(* IEC 61131-3 sources: SortJet_MasterSPS_Aufbau.fbsproj/09_Station/Shuttle/[101,102] Shuttle/Aktionen, 4 files *)

(* ---- Shuttle_Ansteuerung_Ressourcen_FB_V01_00_00.fb.st ---- *)
(* METADATA
{
	"v3Meta": {
		"objectGuid": "9404f6fa-2a6f-44db-8f42-3f6f32f76ed1"
	}
}
*)
FUNCTION_BLOCK Shuttle_Ansteuerung_Ressourcen_FB_V01_00_00 EXTENDS Basic_Shuttle_Aktion_FB_V01_00_00
VAR_INPUT

  // GREIFER [Ausbaustufe stStationsAufbau.bGreifer]
  bpGreiferAktiv : BOOL;
  Greifer        : REFERENCE TO Shuttle_Greifer_FB_V01_00_00;

END_VAR
VAR
  tonlTimeout : TON;

  // BOOL
  blMitGreifer : BOOL; // Vorab-Auftrag mit Greiferseite und Greifer vorhanden
  blGlasUeberspringen : BOOL; // Vorab ohne Glasaktion: Eintransport aktiv oder gerade gewesen
END_VAR
//-------------------------------------------------------------------------------------------------
// AKTION ANSTEUERUNG RESOURCEN WAEHREND DER QUERFAHRT
//-------------------------------------------------------------------------------------------------
(* Wichtig:
   - Es handelt isch hier um eine Aktion die waehrend der Shuttlequerfahrt [Verfahrauftrag] abgearbeitet wird.
   - Zu beachten ist das:
     => Wenn der Riemen verfahrern werden soll pruefen ob der autarke Vortransport aktiv ist
     => Aktion laeuft parallel zum Verfahrauftrag der Oberflaeche
*)
IF (  BasisStationsParameter.bVorabKomponentenAnsteuerung[wWand]
     AND bpAutomatikAktiv )
THEN

  // Ausnahmesituation
  IF ( Glastransport.bpFehler ) THEN
    Glastransport.bpVortransport              := FALSE;
    Glastransport.bpVortransportRueck         := FALSE;
    Glastransport.bpStarteVorabPositionierung := FALSE;
    Glastransport.bpStarteVorabPositionierungRueckwaertig := FALSE;
    BasisStationsParameter.wFehlerNummer := Glastransport.wpFehlerNr;
    steplAktion := STEP_900_E;
  END_IF

  IF ( Kippen.bpFehler ) THEN
    Kippen.bpPositionieren := FALSE;
    BasisStationsParameter.wFehlerNummer :=  Kippen.wpFehlerNr;
    steplAktion := STEP_900_E;
  END_IF

  IF ( Wandverstellung.bpFehler ) THEN
    Wandverstellung.bpStartePositionierung := FALSE;
    BasisStationsParameter.wFehlerNummer :=  Wandverstellung.wpFehlerNr;
    steplAktion := STEP_900_E;
  END_IF

  IF ( blMitGreifer AND Greifer.bpFehler ) THEN
    Greifer.bpPositionieren                         := FALSE;
    Greifer.bpStarteVorabPositionierungEintransport := FALSE;
    BasisStationsParameter.awFehlerInformationen    := Greifer.awpFehlerInformationen;
    BasisStationsParameter.awFehlerInformationen[1] := Greifer.wpFehlerKennung;
    BasisStationsParameter.wFehlerNummer            := Greifer.wpFehlerNr;
    steplAktion := STEP_900_E;
  END_IF

  (* Hinweis:
     - Starten der Schrittkette
  *)
  CASE steplAktion OF
    // VORAB KOMPONENTEN ANSTEUERUNG ========================
    STEP_0_E:
      BasisStationsParameter.bVorabKomponentenAnsteuerungAbgeschlossen[wWand] := FALSE;
      tonlTimeout( IN := FALSE );

      blMitGreifer :=     bpGreiferAktiv
                      AND ( BasisStationsParameter.pVorAbAuftragsdaten[wWand].stAuftragsOptionen.eGreiferTyp <> eGreiferDefault );

      IF ( BasisStationsParameter.stMKs.stStationsOptionen.bVorAbKomponentenAnsteuerung ) THEN
        steplAktion := STEP_10_E;
      ELSE
        steplAktion := STEP_1000_E;
      END_IF

    // VORAB KOMPONENTEN ANSTEUERUNG WAND 1 ========================
    STEP_10_E:
      (* Hinweis:
         - Wandverstellung ansteuern
         - Kippen ansteuern
         - Erst wenn der Glastransport seinen Eintransport beendet hat: Ein vorzeitig quittierter
           Eintransport (letzte Scheibe, Freigabe Querfahrt) laeuft im Glastransport noch weiter,
           waehrend bEintransport bereits FALSE ist. Kippen, Wandverstellung und Greifer duerfen
           die noch fahrende Scheibe nicht beeinflussen (Fehler: Scheibe faehrt auf den Auslaufstopp).
      *)
      IF (     NOT Glastransport.bpEintransport
           AND NOT Glastransport.bpRueckwaertsEintransportieren )
      THEN
        Wandverstellung.epSollStellung         := BasisStationsParameter.pVorAbAuftragsdaten[wWand].stAuftragsOptionen.eDickenverstellung;
        Wandverstellung.bpStartePositionierung := TRUE;

        IF BasisStationsParameter.pVorAbAuftragsdaten[wWand].stAuftragsOptionen.eKippen_SollPosition <> eKippen_Default THEN
          Kippen.epZielPosition := BasisStationsParameter.pVorAbAuftragsdaten[wWand].stAuftragsOptionen.eKippen_SollPosition;
          Kippen.bpPositionieren := TRUE;
        END_IF

        steplAktion := STEP_20_E;
      END_IF

    // VORAB KOMPONENTEN ANSTEUERUNG WAND 1 ========================
    STEP_20_E:
      (* Hinweis:
         - Glastransport ansteuern
         - Laeuft der Eintransport noch (bEintransport) oder ist er gerade abgeschlossen (Eintransport gewesen),
           liegt die Scheibe definiert: die Glasaktion der Vorab entfaellt, es wird nicht gewartet
         - Jede weitere Vorab positioniert die Scheibe neu (Sensor erst freifahren, dann neu anfahren)
      *)
      blGlasUeberspringen := BasisStationsParameter.bEintransport[wWand]
                             OR BasisStationsParameter.bEintransportGewesen[wWand];
      BasisStationsParameter.bEintransportGewesen[wWand] := FALSE;

      IF ( NOT blGlasUeberspringen
           AND NOT Glastransport.bpEintransport
           AND NOT Glastransport.bpRueckwaertsEintransportieren )
      THEN

        CASE BasisStationsParameter.pVorAbAuftragsdaten[wWand].stAuftragsOptionen.eGlastransport OF

          eGlastransport_Default:
            ;

          eGlastransport_AufEinlauf:
            Glastransport.bpStarteVorabPositionierungRueckwaertig := NOT Glastransport.bpAuftragAktiv;

          eGlastransport_AufEinlaufVorab:
            Glastransport.bpVortransportRueck := TRUE;

          eGlastransport_AufAuslauf,
            eGlastransport_AufAuslaufVorab:
            Glastransport.bpStarteVorabPositionierung := NOT Glastransport.bpAuftragAktiv;

        END_CASE

      END_IF

      (* Hinweis:
         - Greifer [Ausbaustufe] waehrend der Querfahrt vorpositionieren
           => Austransport: Greifer hinter die Glaskante stellen
           => Eintransport: Greifer an die Wandseite stellen und ausfahren
         - Entfaellt solange der Eintransport noch aktiv ist (Auftrag oder Glastransport)
      *)
      IF (     blMitGreifer
           AND NOT Greifer.bpAuftragAktiv
           AND NOT BasisStationsParameter.bEintransport[wWand]
           AND NOT Glastransport.bpEintransport
           AND NOT Glastransport.bpRueckwaertsEintransportieren )
      THEN
        Greifer.epGreiferTyp := BasisStationsParameter.pVorAbAuftragsdaten[wWand].stAuftragsOptionen.eGreiferTyp;

        IF ( BasisStationsParameter.pVorAbAuftragsdaten[wWand].wAuftragstyp.0 ) THEN
          Greifer.rpGlaslaenge    := BasisStationsParameter.pVorAbAuftragsdaten[wWand].rLaenge;
          Greifer.bpPositionieren := TRUE;
        ELSE
          Greifer.bpStarteVorabPositionierungEintransport := NOT Greifer.bpVorpositioniertEintransport;
        END_IF
      END_IF

      tonlTimeout( IN := FALSE );
      steplAktion := STEP_100_E;

    // VORAB KOMPONENTEN ANSTEUERUNG WAND 1 ========================
    STEP_100_E:
      (* Hinweis:
         - Einsammeln aller ausgelösten Ereignisse auf bpDone
      *)
      // Nach 60s Fehler melden, dass die Komponenten nicht fertig werden
      tonlTimeout(IN := TRUE, PT := T#60S);

      IF (   ( Kippen.bpDone OR NOT Kippen.bpPositionieren )
           AND (( Glastransport.bpVortransport AND Glastransport.bpDone) OR NOT Glastransport.bpVortransport)
           AND (( Glastransport.bpVortransportRueck AND Glastransport.bpDone) OR NOT Glastransport.bpVortransportRueck)
           AND (( Glastransport.bpStarteVorabPositionierung AND Glastransport.bpDone) OR NOT Glastransport.bpStarteVorabPositionierung)
           AND (( Glastransport.bpStarteVorabPositionierungRueckwaertig AND Glastransport.bpDone) OR NOT Glastransport.bpStarteVorabPositionierungRueckwaertig)
           AND (( Wandverstellung.bpStartePositionierung AND Wandverstellung.bpDone) OR NOT Wandverstellung.bpStartePositionierung)
           AND (    NOT blMitGreifer
                 OR (     (( Greifer.bpPositionieren AND Greifer.bpPositionierungAbgeschlossen ) OR NOT Greifer.bpPositionieren )
                      AND (( Greifer.bpStarteVorabPositionierungEintransport AND Greifer.bpVorabPositionierungEintransportAbgeschlossen ) OR NOT Greifer.bpStarteVorabPositionierungEintransport ) ) ) )
      THEN

        Glastransport.bpVortransport                    := FALSE;
        Glastransport.bpVortransportRueck               := FALSE;
        Glastransport.bpStarteVorabPositionierung       := FALSE;
        Glastransport.bpStarteVorabPositionierungRueckwaertig := FALSE;

        Wandverstellung.bpStartePositionierung          := FALSE;
        Kippen.bpPositionieren                          := FALSE;

        IF ( blMitGreifer ) THEN
          Greifer.bpPositionieren                         := FALSE;
          Greifer.bpStarteVorabPositionierungEintransport := FALSE;
        END_IF

        steplAktion := STEP_1000_E;
      END_IF

      IF tonlTimeout.Q THEN
        BasisStationsParameter.wFehlerNummer := cMELDUNG_STATION_VORABKOMPONENTENANSTEUERUN_NOT_DONE;
        steplAktion := STEP_900_E;
      END_IF

    // VORAB KOMPONENTEN ANSTEUERUNG WAND 1 ========================
    STEP_900_E:
      BasisStationsParameter.bFehler := TRUE;

    // VORAB KOMPONENTEN ANSTEUERUNG WAND 1 ========================
    STEP_1000_E:

      Glastransport.bpVortransport                    := FALSE;
      Glastransport.bpVortransportRueck               := FALSE;
      Glastransport.bpStarteVorabPositionierung       := FALSE;
      Glastransport.bpStarteVorabPositionierungRueckwaertig := FALSE;

      Wandverstellung.bpStartePositionierung          := FALSE;
      Kippen.bpPositionieren                          := FALSE;

      BasisStationsParameter.bVorabKomponentenAnsteuerungAbgeschlossen[wWand] := TRUE;

  // VORAB KOMPONENTEN ANSTEUERUNG WAND 1 ========================
  END_CASE

END_IF

IF ( NOT BasisStationsParameter.bVorabKomponentenAnsteuerung[wWand] ) THEN

  IF ( steplAktion > STEP_0_E ) THEN

    IF ( NOT BasisStationsParameter.bVorabKomponentenAnsteuerungAbgeschlossen[wWand] ) THEN

      Glastransport.bpVortransport                    := FALSE;
      Glastransport.bpVortransportRueck               := FALSE;
      Glastransport.bpStarteVorabPositionierung       := FALSE;
      Glastransport.bpStarteVorabPositionierungRueckwaertig := FALSE;

      Wandverstellung.bpStartePositionierung          := FALSE;
      Kippen.bpPositionieren                                   := FALSE;
    END_IF

    IF ( blMitGreifer ) THEN
      Greifer.bpPositionieren                         := FALSE;
      Greifer.bpStarteVorabPositionierungEintransport := FALSE;
      blMitGreifer := FALSE;
    END_IF

    BasisStationsParameter.bVorabKomponentenAnsteuerungAbgeschlossen[wWand] := FALSE;

    steplAktion := STEP_0_E;
  END_IF

END_IF
END_FUNCTION_BLOCK

(* ---- Shuttle_Austransport_FB_V01_00_00.fb.st ---- *)
(* METADATA
{
	"v3Meta": {
		"objectGuid": "aea75a09-065c-4155-9284-9233b13eb99a"
	}
}
*)
FUNCTION_BLOCK Shuttle_Austransport_FB_V01_00_00 EXTENDS Basic_Shuttle_Aktion_FB_V01_00_00
VAR_INPUT

  // GREIFER [Ausbaustufe stStationsAufbau.bGreifer]
  bpGreiferAktiv : BOOL;
  Greifer        : REFERENCE TO Shuttle_Greifer_FB_V01_00_00;

END_VAR
VAR

  // BOOL
  blMitGreifer : BOOL; // Austransport mit dem Greifer (Greifer vorhanden und Greiferseite im Auftrag)

  // TIMER
  tonlUeberwachungGreifer : TON;

END_VAR
VAR CONSTANT

  // TIME
  cZEIT_UEBERWACHUNG_GREIFER : TIME := T#120S; // Gesamtueberwachung je Greifer-Schritt (die Wartestellen ueberwacht der Greifer selbst)

END_VAR
//-------------------------------------------------------------------------------------------------
// AKTION AUSTRANSPORT WAND 1
//-------------------------------------------------------------------------------------------------
(* Hinweis:
   - Es handelt sich hier um einen Austransport in einen Faecherwagen
*)
IF (  BasisStationsParameter.bAustransport[wWand]
     AND bpAutomatikAktiv )
THEN

  // Ausnahmesituation
  IF ( Glastransport.bpFehler ) THEN
    Glastransport.bpAustransport := FALSE;
    BasisStationsParameter.wFehlerNummer :=  Glastransport.wpFehlerNr;
    steplAktion := STEP_900_E;
  END_IF

  IF ( Kippen.bpFehler ) THEN
    Kippen.bpPositionieren := FALSE;
    BasisStationsParameter.wFehlerNummer :=  Kippen.wpFehlerNr;
    steplAktion := STEP_900_E;
  END_IF

  IF ( Wandverstellung.bpFehler ) THEN
    Wandverstellung.bpStartePositionierung := FALSE;
    BasisStationsParameter.wFehlerNummer :=  Wandverstellung.wpFehlerNr;
    steplAktion := STEP_900_E;
  END_IF

  IF ( Geblaese.bpFehler ) THEN
    BasisStationsParameter.wFehlerNummer := cMELDUNG_ANTRIEB_GEBLAESE;
    steplAktion:=STEP_900_E;
  END_IF

  IF ( blMitGreifer AND Greifer.bpFehler ) THEN
    Greifer.bpPositionieren                       := FALSE;
    Greifer.bpStarteAustransport                  := FALSE;
    Glastransport.bpStarteGlasPositionierungGreifer := FALSE;
    Glastransport.bpStarteKorrekturfahrt          := FALSE;
    BasisStationsParameter.awFehlerInformationen  := Greifer.awpFehlerInformationen;
    BasisStationsParameter.awFehlerInformationen[1] := Greifer.wpFehlerKennung;
    BasisStationsParameter.wFehlerNummer          := Greifer.wpFehlerNr;
    steplAktion := STEP_900_E;
  END_IF

  CASE steplAktion OF
    // AUSTRANSPORT =====================================
    STEP_0_E:
      (* Hinweis:
         - Variablen zuruecksetzen
      *)
      BasisStationsParameter.bAustransportAbgeschlossen[wWand]    := FALSE;

      blMitGreifer :=     bpGreiferAktiv
                      AND ( BasisStationsParameter.pAuftrag[wWand].stAuftragsOptionen.eGreiferTyp <> eGreiferDefault );

      steplAktion := STEP_10_E;

    // AUSTRANSPORT =====================================
    STEP_10_E:
      (* Hinweis:
         - Pruefen ob die Zielposition erreicht wurde
      *)
      IF ( bpZielPositionErreicht ) THEN
        steplAktion := STEP_20_E;

      ELSE
        BasisStationsParameter.awFehlerInformationen[1] := REAL_TO_WORD(BasisStationsParameter.rAktuellePositionQuerfahrt);
        BasisStationsParameter.awFehlerInformationen[2] := REAL_TO_WORD(BasisStationsParameter.pAuftrag[wWand].rVorabPosition);
        BasisStationsParameter.wFehlerNummer := cMELDUNG_QUERFAHRT_SOLLPOSITION_NICHT_ERREICHT;

        steplAktion := STEP_900_E;

      END_IF

    // AUSTRANSPORT =====================================
    STEP_20_E:
      // ---------------------------------------------------------------------------------------
      //  ANSTEUERUNG KOMPONENTEN
      //
      //  Hinweis:
      //  - Sicherstellen dass das Geblaese aktiv  und keine Vorab- Auftrag aktiv sind
      // ---------------------------------------------------------------------------------------

      IF (  bpGeblaeseAktiv
           AND NOT bpVorAbAuftragAktiv )
      THEN

        (* Hinweis:
           - Anstellen der Dicken-/ Wandverstellung in Abhängigkeit der Glasdicke
        *)
        Wandverstellung.epSollStellung         := BasisStationsParameter.pAuftrag[wWand].stAuftragsOptionen.eDickenverstellung;
        Wandverstellung.bpStartePositionierung := FALSE;

        (* Hinweis:
           - Shuttle in die passende Position kippen
        *)
        Kippen.epZielPosition := BasisStationsParameter.pAuftrag[wWand].stAuftragsOptionen.eKippen_SollPosition;
        Kippen.bpPositionieren := TRUE;

        steplAktion := STEP_30_E;

      END_IF

      (* Fehlerbehandlung:
         - Geblaese
      *)
      IF ( Geblaese.bpFehler ) THEN
        BasisStationsParameter.wFehlerNummer := cMELDUNG_ANTRIEB_GEBLAESE;
        steplAktion := STEP_900_E;
      END_IF

    // AUSTRANSPORT =====================================
    STEP_30_E:
      (* Hinweis:
         - Wandverstellung gefahren ?
      *)
      IF ( (  Wandverstellung.bpDone OR  NOT Wandverstellung.bpStartePositionierung )
           AND (  Kippen.bpDone OR NOT Kippen.bpPositionieren ) )
      THEN
        Kippen.bpPositionieren := FALSE;

        Wandverstellung.bpStartePositionierung := FALSE;

        IF ( blMitGreifer ) THEN
          steplAktion := STEP_200_E;
        ELSE
          steplAktion := STEP_100_E;
        END_IF
      END_IF

      // Ausnahmesituation
      //   - Komponenten
      IF ( Wandverstellung.bpFehler ) THEN
        Wandverstellung.bpStartePositionierung := FALSE;
        BasisStationsParameter.wFehlerNummer :=  Wandverstellung.wpFehlerNr;
        steplAktion := STEP_900_E;
      END_IF

    // AUSTRANSPORT =====================================
    STEP_50_E:
      (* Hinweis:
         - Kippvorgang beendet
         - Vortransport beendet
           WICHTIG:
         - Wenn der Empfaenger eine Station ist kann der Vortransport abgebrochen werden
      *)
      IF ( Glastransport.bpDone
           OR BasisStationsParameter.InGlasTransportNachfolger[wWand].bBereitZumEintransport )
      THEN

        Glastransport.bpVortransport      := FALSE;
        Glastransport.bpVortransportRueck := FALSE;

        steplAktion := STEP_100_E;
      END_IF

    // AUSTRANSPORT =====================================
    STEP_100_E:
      // ---------------------------------------------------------------------------------------
      //  STARTEN DES AUSTRANSPORTS
      //
      //  Hinweis:
      //  - Unterscheidung ob Rueckwertiger- Transport
      // ---------------------------------------------------------------------------------------
      (* Hinweis:
         - Ein vorzeitig quittierter Eintransport laeuft im Glastransport selbststaendig zu Ende und wird nicht abgebrochen
         - Der Austransport startet erst danach (Ueberwachung durch die Eintransport-Kette selbst)
      *)
      IF ( NOT Glastransport.bpEintransport
           AND NOT Glastransport.bpRueckwaertsEintransportieren )
      THEN
        Glastransport.pAuftrag := BasisStationsParameter.pAuftrag[wWand];

        Glastransport.bpAustransport                 := NOT BasisStationsParameter.bRueckwaertsTransportieren[wWand];
        Glastransport.bpRueckwaertsAustransportieren := BasisStationsParameter.bRueckwaertsTransportieren[wWand];

        steplAktion := STEP_110_E;
      END_IF

    // AUSTRANSPORT ==============================
    STEP_110_E:
      (* Hinweis:
         - Scheibenzaehlen waerend der Glastransport arbeitet.
            Verarbeitung im ShuttleJobs Baustein
      *)
      bprtScheibe := Glastransport.bprtScheibe;

      (* Hinweis [Glastransport]:
         - Austransport der Scheiben abgeschlossen
      *)
      IF ( Glastransport.bpDone ) THEN
        Glastransport.bpAustransport                  := FALSE;
        Glastransport.bpRueckwaertsAustransportieren  := FALSE;
        steplAktion := STEP_1000_E;
      END_IF

    // AUSTRANSPORT GREIFER ======================
    STEP_200_E:
      // ---------------------------------------------------------------------------------------
      //  AUSTRANSPORT MIT DEM GREIFER [AUSBAUSTUFE]
      //
      //  Hinweis:
      //  - Keine Vorab-Ansteuerung und kein anderer Ablauf des Greifers aktiv
      //  - Scheibe ueber den Sensor der Greiferseite positionieren und den Greifer hinter die Glaskante stellen
      // ---------------------------------------------------------------------------------------
      tonlUeberwachungGreifer( IN := TRUE, PT := cZEIT_UEBERWACHUNG_GREIFER );

      IF (     NOT bpVorAbAuftragAktiv
           AND NOT Greifer.bpAuftragAktiv )
      THEN
        tonlUeberwachungGreifer( IN := FALSE );

        Greifer.epGreiferTyp    := BasisStationsParameter.pAuftrag[wWand].stAuftragsOptionen.eGreiferTyp;
        Greifer.pAuftrag        := BasisStationsParameter.pAuftrag[wWand];
        Greifer.rpGlaslaenge    := BasisStationsParameter.pAuftrag[wWand].rAuftragsLaenge;
        Greifer.bpPositionieren := TRUE;

        Glastransport.pAuftrag                          := BasisStationsParameter.pAuftrag[wWand];
        Glastransport.bpGlasPositionierungEinlaufseite  := ( BasisStationsParameter.pAuftrag[wWand].stAuftragsOptionen.eGreiferTyp = eGreiferEinlaufseite );
        Glastransport.rpWegGlasUebergabeposition        := Greifer.rpWegGlasUebergabeposition;
        Glastransport.bpStarteGlasPositionierungGreifer := TRUE;

        steplAktion := STEP_210_E;
      END_IF

      IF ( tonlUeberwachungGreifer.Q ) THEN
        tonlUeberwachungGreifer( IN := FALSE );
        BasisStationsParameter.wFehlerNummer := cMELDUNG_GREIFER_STOESSEL_ABLAUF_ZEITUEBERSCHREITUNG;
        steplAktion := STEP_900_E;
      END_IF

    // AUSTRANSPORT GREIFER ======================
    STEP_210_E:
      (* Hinweis:
         - Weg ueber den Sensor laufend aus dem Greifer uebernehmen (Auftragsdaten im Greifer aktualisiert)
         - Scheibe und Greifer positioniert
      *)
      Glastransport.rpWegGlasUebergabeposition := Greifer.rpWegGlasUebergabeposition;

      tonlUeberwachungGreifer( IN := TRUE, PT := cZEIT_UEBERWACHUNG_GREIFER );

      IF (     Glastransport.bpGlasPositionierungGreiferAbgeschlossen
           AND Greifer.bpPositionierungAbgeschlossen )
      THEN
        tonlUeberwachungGreifer( IN := FALSE );
        Glastransport.bpStarteGlasPositionierungGreifer := FALSE;
        Greifer.bpPositionieren := FALSE;
        steplAktion := STEP_220_E;
      END_IF

      IF ( tonlUeberwachungGreifer.Q ) THEN
        tonlUeberwachungGreifer( IN := FALSE );
        Glastransport.bpStarteGlasPositionierungGreifer := FALSE;
        Greifer.bpPositionieren := FALSE;
        BasisStationsParameter.wFehlerNummer := cMELDUNG_GREIFER_STOESSEL_ABLAUF_ZEITUEBERSCHREITUNG;
        steplAktion := STEP_900_E;
      END_IF

    // AUSTRANSPORT GREIFER ======================
    STEP_220_E:
      (* Hinweis:
         - Austransport mit dem Greifer starten
      *)
      Greifer.bpStarteAustransport := TRUE;
      steplAktion := STEP_230_E;

    // AUSTRANSPORT GREIFER ======================
    STEP_230_E:
      (* Hinweis:
         - Quittierung der Scheibe
         - Austransport mit dem Greifer abgeschlossen
      *)
      bprtScheibe := Greifer.bprtScheibe;

      tonlUeberwachungGreifer( IN := TRUE, PT := cZEIT_UEBERWACHUNG_GREIFER );

      IF ( Greifer.bpAustransportAbgeschlossen ) THEN
        tonlUeberwachungGreifer( IN := FALSE );
        Greifer.bpStarteAustransport := FALSE;
        steplAktion := STEP_240_E;
      END_IF

      IF ( tonlUeberwachungGreifer.Q ) THEN
        tonlUeberwachungGreifer( IN := FALSE );
        Greifer.bpStarteAustransport := FALSE;
        BasisStationsParameter.wFehlerNummer := cMELDUNG_GREIFER_STOESSEL_ABLAUF_ZEITUEBERSCHREITUNG;
        steplAktion := STEP_900_E;
      END_IF

    // AUSTRANSPORT GREIFER ======================
    STEP_240_E:
      (* Hinweis:
         - Korrekturfahrt des Glastransports: Sensor der Greiferseite frei fahren
      *)
      bprtScheibe := FALSE;

      Glastransport.bpKorrekturfahrtRueckwaerts := ( BasisStationsParameter.pAuftrag[wWand].stAuftragsOptionen.eGreiferTyp = eGreiferAuslaufseite );
      Glastransport.bpStarteKorrekturfahrt      := TRUE;

      steplAktion := STEP_250_E;

    // AUSTRANSPORT GREIFER ======================
    STEP_250_E:
      tonlUeberwachungGreifer( IN := TRUE, PT := cZEIT_UEBERWACHUNG_GREIFER );

      IF ( Glastransport.bpKorrekturfahrtAbgeschlossen ) THEN
        tonlUeberwachungGreifer( IN := FALSE );
        Glastransport.bpStarteKorrekturfahrt := FALSE;
        steplAktion := STEP_1000_E;
      END_IF

      IF ( tonlUeberwachungGreifer.Q ) THEN
        tonlUeberwachungGreifer( IN := FALSE );
        Glastransport.bpStarteKorrekturfahrt := FALSE;
        BasisStationsParameter.wFehlerNummer := cMELDUNG_GREIFER_STOESSEL_ABLAUF_ZEITUEBERSCHREITUNG;
        steplAktion := STEP_900_E;
      END_IF

    // AUSTRANSPORT ==============================
    STEP_900_E:
      Glastransport.bpAustransport                 := FALSE;
      Glastransport.bpRueckwaertsAustransportieren := FALSE;

      Glastransport.bpVortransport      := FALSE;
      Glastransport.bpVortransportRueck := FALSE;

      BasisStationsParameter.bFehler := TRUE;

    // AUSTRANSPORT ==============================
    STEP_1000_E:
      BasisStationsParameter.bAustransportAbgeschlossen[wWand] := TRUE;

  // AUSTRANSPORT ==============================
  END_CASE
ELSE

  IF ( steplAktion > STEP_0_E ) THEN

    (* Hinweis:
       - Zuruecksetzen
    *)
    IF ( NOT BasisStationsParameter.bAustransportAbgeschlossen[wWand] ) THEN
      Kippen.bpPositionieren := FALSE;

      Wandverstellung.bpStartePositionierung := FALSE;

    END_IF

    bprtScheibe := FALSE;

    BasisStationsParameter.bAustransportAbgeschlossen[wWand] := FALSE;

    Glastransport.bpAustransport                 := FALSE;
    Glastransport.bpRueckwaertsAustransportieren := FALSE;

    Glastransport.bpVortransport          := FALSE;
    Glastransport.bpVortransportRueck     := FALSE;

    IF ( blMitGreifer ) THEN
      Greifer.bpPositionieren                         := FALSE;
      Greifer.bpStarteAustransport                    := FALSE;
      Glastransport.bpStarteGlasPositionierungGreifer := FALSE;
      Glastransport.bpStarteKorrekturfahrt            := FALSE;
      tonlUeberwachungGreifer( IN := FALSE );
      blMitGreifer := FALSE;
    END_IF

    steplAktion := STEP_0_E;

  END_IF

END_IF
END_FUNCTION_BLOCK

(* ---- Shuttle_Durchtransport_FB_V01_00_00.fb.st ---- *)
(* METADATA
{
	"v3Meta": {
		"objectGuid": "fde90b53-97e1-44a2-93b0-a69a2d65f26b"
	}
}
*)
FUNCTION_BLOCK Shuttle_Durchtransport_FB_V01_00_00 EXTENDS Basic_Shuttle_Aktion_FB_V01_00_00
VAR
END_VAR
//-------------------------------------------------------------------------------------------------
// DURCHTRANSPORT WAND 1
//-------------------------------------------------------------------------------------------------
IF ( BasisStationsParameter.bDurchtransport[wWand]
     AND bpAutomatikAktiv )
THEN

  // Ausnahmesituation
  IF ( Glastransport.bpFehler ) THEN
    Glastransport.bpDurchtransport := FALSE;
    BasisStationsParameter.wFehlerNummer :=  Glastransport.wpFehlerNr;
    steplAktion := STEP_900_E;
  END_IF

  IF ( Kippen.bpFehler ) THEN
    Kippen.bpPositionieren := FALSE;
    BasisStationsParameter.wFehlerNummer :=  Kippen.wpFehlerNr;
    steplAktion := STEP_900_E;
  END_IF

  IF ( Wandverstellung.bpFehler ) THEN
    Wandverstellung.bpStartePositionierung := FALSE;
    BasisStationsParameter.wFehlerNummer :=  Wandverstellung.wpFehlerNr;
    steplAktion := STEP_900_E;
  END_IF

  IF ( Geblaese.bpFehler ) THEN
    BasisStationsParameter.wFehlerNummer := cMELDUNG_ANTRIEB_GEBLAESE;
    steplAktion:=STEP_900_E;
  END_IF

  CASE steplAktion OF
    // DURCHTRANSPORT ==============================
    STEP_0_E:
      (* Hinweis:
         - Variablen zuruecksetzen
      *)
      BasisStationsParameter.bEintransportAbgeschlossen[wWand] := FALSE;

      steplAktion := STEP_10_E;

    // DURCHTRANSPORT ==============================
    STEP_10_E:
      (* Hinweis:
         - Pruefen ob die Geblase aktiv sind
         - Quellstation pruefen
      *)
      IF ( bpGeblaeseAktiv ) THEN

        IF ( NOT bpVorAbAuftragAktiv ) THEN

          (* Hinweis:
             - Anstellen der Dicken-/ Wandverstellung in Abhängigkeit der Glasdicke
          *)
          Wandverstellung.epSollStellung         := BasisStationsParameter.pAuftrag[wWand].stAuftragsOptionen.eDickenverstellung;
          Wandverstellung.bpStartePositionierung := TRUE;

          Kippen.epZielPosition := BasisStationsParameter.pAuftrag[wWand].stAuftragsOptionen.eKippen_SollPosition;
          Kippen.bpPositionieren := TRUE;

          steplAktion := STEP_20_E;
        END_IF

      END_IF

    // DURCHTRANSPORT ==============================
    STEP_20_E:
      // Verfahrauftrag ans Shuttle uebergeben [Verfahrueberwachung]:
      //   - Pruefen ob das Shuttel zum verfahren freigegeben ist, wenn ja Zielposition
      //     aus dem Auftrag uebergeben.
      IF ( bpZielPositionErreicht ) THEN
        steplAktion := STEP_30_E;

      ELSE
        BasisStationsParameter.awFehlerInformationen[1] := REAL_TO_WORD(BasisStationsParameter.rAktuellePositionQuerfahrt);
        BasisStationsParameter.awFehlerInformationen[2] := REAL_TO_WORD(BasisStationsParameter.pAuftrag[wWand].rVorabPosition);
        BasisStationsParameter.wFehlerNummer := cMELDUNG_QUERFAHRT_SOLLPOSITION_NICHT_ERREICHT;

        steplAktion := STEP_900_E;
      END_IF

    // DURCHTRANSPORT ==============================
    STEP_30_E:
      (* Hinweis:
         - Sicherstellen das die Wand auch wirklich ihre Soll-Position erreicht hat
      *)
      Wandverstellung.epSollStellung         := BasisStationsParameter.pAuftrag[wWand].stAuftragsOptionen.eDickenverstellung;
      Wandverstellung.bpStartePositionierung := TRUE;

      (* Hinweis:
         - Dickenverstellung-Abschluss
      *)
      IF Wandverstellung.bpDone THEN
        Wandverstellung.bpStartePositionierung := FALSE;
        steplAktion := STEP_40_E;
      END_IF

    // DURCHTRANSPORT ==============================
    STEP_40_E:
      // ---------------------------------------------------------------------------------------
      //  KIPP- VORGANG ABSCHLIESSEN
      //
      //  Hinweis:
      //  - n/c
      // ---------------------------------------------------------------------------------------

      IF ( Kippen.bpDone OR NOT Kippen.bpPositionieren )
         AND ( Kippen.epKippStatus = BasisStationsParameter.pAuftrag[wWand].stAuftragsOptionen.eKippen_SollPosition)
      THEN
        Kippen.bpPositionieren  := FALSE;
        steplAktion := STEP_100_E;
      END_IF

    // DURCHTRANSPORT ==============================
    STEP_100_E:
      // ---------------------------------------------------------------------------------------
      //  STARTEN DES DURCHTRANSPORTS
      // ---------------------------------------------------------------------------------------

      Glastransport.pAuftrag := BasisStationsParameter.pAuftrag[wWand];
      Glastransport.bpDurchtransport := TRUE;

      steplAktion := STEP_110_E;

    // DURCHTRANSPORT ==============================
    STEP_110_E:
      (* Hinweis:
         - Quittierung der Scheibe
      *)
      bprtScheibe := Glastransport.bprtScheibe;

      (* Hinweis:
         - Eintransport der Scheiben abgeschlossen
      *)
      IF ( Glastransport.bpDone ) THEN
        Glastransport.bpDurchtransport := FALSE;
        steplAktion := STEP_200_E;
      END_IF

    // DURCHTRANSPORT ==============================
    STEP_200_E:
      (* Hinweis:
         - Kippen ansteuern
      *)
      bprtScheibe := Glastransport.bprtScheibe;

      Kippen.epZielPosition := BasisStationsParameter.pAuftrag[wWand].stAuftragsOptionen.eKippen_SollPosition_NachAustransport;
      Kippen.bpPositionieren := TRUE;

      steplAktion := STEP_210_E;

    // DURCHTRANSPORT ==============================
    STEP_210_E:
      (* Hinweis:
         - Quittierung der Scheibe
      *)
      bprtScheibe := Glastransport.bprtScheibe;

      (* Hinweis:
         - Kippen abschließen
      *)
      IF Kippen.bpDone THEN
        Kippen.bpPositionieren := FALSE;
        steplAktion := STEP_1000_E;
      END_IF

    // DURCHTRANSPORT ==============================
    STEP_900_E:
      BasisStationsParameter.bFehler := TRUE;

    // DURCHTRANSPORT ==============================
    STEP_1000_E:
      bprtScheibe := FALSE;
      BasisStationsParameter.bDurchtransportAbgeschlossen[wWand] := TRUE;

  // DURCHTRANSPORT ==============================
  END_CASE
ELSE

  IF (steplAktion > STEP_0_E) THEN

    BasisStationsParameter.bDurchtransportAbgeschlossen[wWand] := FALSE;
    bprtScheibe := FALSE;

    Glastransport.bpDurchtransport := FALSE;

    Kippen.bpPositionieren := FALSE;
    Wandverstellung.bpStartePositionierung := FALSE;

    steplAktion := STEP_0_E;
  END_IF

END_IF
END_FUNCTION_BLOCK

(* ---- Shuttle_Eintransport_FB_V01_00_00.fb.st ---- *)
(* METADATA
{
	"v3Meta": {
		"objectGuid": "658aa591-8bd2-427d-a42c-c4e6e57fe5c7"
	}
}
*)
FUNCTION_BLOCK Shuttle_Eintransport_FB_V01_00_00 EXTENDS Basic_Shuttle_Aktion_FB_V01_00_00
VAR_INPUT

  // GREIFER [Ausbaustufe stStationsAufbau.bGreifer]
  bpGreiferAktiv : BOOL;
  Greifer        : REFERENCE TO Shuttle_Greifer_FB_V01_00_00;

END_VAR
VAR

  // BOOL
  blMitGreifer : BOOL; // Eintransport mit dem Greifer (Greifer vorhanden und Greiferseite im Auftrag)

  // TIMER
  tonlUeberwachungGreifer : TON;

END_VAR
VAR CONSTANT

  // TIME
  cZEIT_UEBERWACHUNG_GREIFER : TIME := T#120S; // Gesamtueberwachung je Greifer-Schritt (die Wartestellen ueberwacht der Greifer selbst)

END_VAR
//-------------------------------------------------------------------------------------------------
// EINTRANSPORT WAND 1
//-------------------------------------------------------------------------------------------------
IF ( BasisStationsParameter.bEintransport[wWand]
     AND bpAutomatikAktiv )
THEN

  // Ausnahmesituation
  IF ( Glastransport.bpFehler ) THEN
    Glastransport.bpEintransport := FALSE;
    BasisStationsParameter.wFehlerNummer :=  Glastransport.wpFehlerNr;
    steplAktion := STEP_900_E;
  END_IF

  IF ( Kippen.bpFehler ) THEN
    Kippen.bpPositionieren := FALSE;
    BasisStationsParameter.wFehlerNummer :=  Kippen.wpFehlerNr;
    steplAktion := STEP_900_E;
  END_IF

  IF ( Wandverstellung.bpFehler ) THEN
    Wandverstellung.bpStartePositionierung := FALSE;
    BasisStationsParameter.wFehlerNummer :=  Wandverstellung.wpFehlerNr;
    steplAktion := STEP_900_E;
  END_IF

  IF ( Geblaese.bpFehler ) THEN
    BasisStationsParameter.wFehlerNummer := cMELDUNG_ANTRIEB_GEBLAESE;
    steplAktion:=STEP_900_E;
  END_IF

  IF ( blMitGreifer AND Greifer.bpFehler ) THEN
    Greifer.bpStarteVorabPositionierungEintransport := FALSE;
    Greifer.bpStarteEintransport                    := FALSE;
    Glastransport.bpStarteKorrekturfahrt            := FALSE;
    BasisStationsParameter.awFehlerInformationen    := Greifer.awpFehlerInformationen;
    BasisStationsParameter.awFehlerInformationen[1] := Greifer.wpFehlerKennung;
    BasisStationsParameter.wFehlerNummer            := Greifer.wpFehlerNr;
    steplAktion := STEP_900_E;
  END_IF

  CASE steplAktion OF
    // EINTRANSPORT ==============================
    STEP_0_E:
      (* Hinweis:
         - Variablen zuruecksetzen
      *)
      BasisStationsParameter.bEintransportAbgeschlossen[wWand] := FALSE;

      blMitGreifer :=     bpGreiferAktiv
                      AND ( BasisStationsParameter.pAuftrag[wWand].stAuftragsOptionen.eGreiferTyp <> eGreiferDefault );

      steplAktion := STEP_10_E;

    // EINTRANSPORT ==============================
    STEP_10_E:
      (* Hinweis:
         - Pruefen ob die Geblase aktiv sind
         - Wandverstellung starten
         - Kippen starten
      *)
      IF ( bpGeblaeseAktiv ) THEN

        IF ( NOT bpVorAbAuftragAktiv ) THEN

          Wandverstellung.epSollStellung         := BasisStationsParameter.pAuftrag[wWand].stAuftragsOptionen.eDickenverstellung;
          Wandverstellung.bpStartePositionierung := TRUE;

          Kippen.epZielPosition := BasisStationsParameter.pAuftrag[wWand].stAuftragsOptionen.eKippen_SollPosition;
          Kippen.bpPositionieren := TRUE;

          steplAktion := STEP_20_E;
        END_IF

      END_IF

    // EINTRANSPORT ==============================
    STEP_20_E:
      // Verfahrauftrag ans Shuttle uebergeben [Verfahrueberwachung]:
      //   - Pruefen ob das Shuttel zum verfahren freigegeben ist, wenn ja Zielposition
      //     aus dem Auftrag uebergeben.
      IF ( bpZielPositionErreicht ) THEN
        steplAktion := STEP_30_E;

      ELSE
        BasisStationsParameter.awFehlerInformationen[1] := REAL_TO_WORD(BasisStationsParameter.rAktuellePositionQuerfahrt);
        BasisStationsParameter.awFehlerInformationen[2] := REAL_TO_WORD(BasisStationsParameter.pAuftrag[wWand].rVorabPosition);
        BasisStationsParameter.wFehlerNummer := cMELDUNG_QUERFAHRT_SOLLPOSITION_NICHT_ERREICHT;

        steplAktion := STEP_900_E;
      END_IF

    // EINTRANSPORT ==============================
    STEP_30_E:
      (* Hinweis:
         - Sicherstellen das die Wand auch wirklich ihre Soll-Position erreicht hat
      *)
      Wandverstellung.epSollStellung         := BasisStationsParameter.pAuftrag[wWand].stAuftragsOptionen.eDickenverstellung;
      Wandverstellung.bpStartePositionierung := TRUE;

      (* Hinweis:
         - Dickenverstellung-Abschluss
      *)
      IF Wandverstellung.bpDone THEN
        Wandverstellung.bpStartePositionierung := FALSE;
        steplAktion := STEP_40_E;
      END_IF

    // EINTRANSPORT ==============================
    STEP_40_E:
      (* Hinweis:
         - Kippen abgeschlossen -> pruefen ob Position erreicht
      *)
      IF ( Kippen.bpDone OR NOT Kippen.bpPositionieren )
         AND ( Kippen.epKippStatus = BasisStationsParameter.pAuftrag[wWand].stAuftragsOptionen.eKippen_SollPosition)
      THEN
        Kippen.bpPositionieren  := FALSE;

        IF ( blMitGreifer ) THEN
          steplAktion := STEP_200_E;
        ELSE
          steplAktion := STEP_100_E;
        END_IF
      END_IF

    // EINTRANSPORT ==============================
    STEP_100_E:
      // ---------------------------------------------------------------------------------------
      //  STARTEN DES EINTRANSPORTS
      //
      //  Hinweis:
      //  - Unterscheidung ob Rueckwertiger- Transport
      // ---------------------------------------------------------------------------------------

      Glastransport.bpRueckwaertsEintransportieren   := BasisStationsParameter.bRueckwaertsTransportieren[wWand];
      Glastransport.bpEintransport                   := NOT BasisStationsParameter.bRueckwaertsTransportieren[wWand];

      Glastransport.bpTransferstationTransfershuttle := BasisStationsParameter.bTransferstationTransfershuttle[wWand];
      Glastransport.bpScheibentrennung               := BasisStationsParameter.bScheibentrennen[wWand];
      Glastransport.pAuftrag                         := BasisStationsParameter.pAuftrag[wWand];

      steplAktion := STEP_110_E;

    // EINTRANSPORT ==============================
    STEP_110_E:
      (* Hinweis:
         - Quittierung der Scheibe
      *)
      bprtScheibe := Glastransport.bprtScheibe;

      (* Hinweis:
         - Eintransport der Scheiben abgeschlossen
      *)
      IF ( Glastransport.bpDone ) THEN
        Glastransport.bpEintransport := FALSE;
        Glastransport.bpRueckwaertsEintransportieren := FALSE;
        steplAktion := STEP_1000_E;
      END_IF

      (* Hinweis:
         - Eintransport vorzeitig quittieren damit die Querfahrt starten kann
      *)
      IF (  BasisStationsParameter.pAuftrag[wWand].bLetzteScheibe
           AND Glastransport.bpFreigabeQuerfahrt )
      THEN
        steplAktion := STEP_1000_E;
      END_IF

    // EINTRANSPORT GREIFER ======================
    STEP_200_E:
      // ---------------------------------------------------------------------------------------
      //  EINTRANSPORT MIT DEM GREIFER [AUSBAUSTUFE]
      //
      //  Hinweis:
      //  - Greifer an die Wandseite stellen, sofern er nicht schon vorpositioniert ist
      // ---------------------------------------------------------------------------------------
      Greifer.epGreiferTyp := BasisStationsParameter.pAuftrag[wWand].stAuftragsOptionen.eGreiferTyp;
      Greifer.pAuftrag     := BasisStationsParameter.pAuftrag[wWand];

      Greifer.bpStarteVorabPositionierungEintransport := NOT Greifer.bpVorpositioniertEintransport;

      steplAktion := STEP_210_E;

    // EINTRANSPORT GREIFER ======================
    STEP_210_E:
      (* Hinweis:
         - Greifer vorpositioniert, Eintransport mit dem Greifer starten
      *)
      tonlUeberwachungGreifer( IN := TRUE, PT := cZEIT_UEBERWACHUNG_GREIFER );

      IF (    Greifer.bpVorabPositionierungEintransportAbgeschlossen
           OR Greifer.bpVorpositioniertEintransport )
      THEN
        tonlUeberwachungGreifer( IN := FALSE );
        Greifer.bpStarteVorabPositionierungEintransport := FALSE;
        Greifer.bpStarteEintransport := TRUE;
        steplAktion := STEP_220_E;
      END_IF

      IF ( tonlUeberwachungGreifer.Q ) THEN
        tonlUeberwachungGreifer( IN := FALSE );
        Greifer.bpStarteVorabPositionierungEintransport := FALSE;
        BasisStationsParameter.wFehlerNummer := cMELDUNG_GREIFER_STOESSEL_ABLAUF_ZEITUEBERSCHREITUNG;
        steplAktion := STEP_900_E;
      END_IF

    // EINTRANSPORT GREIFER ======================
    STEP_220_E:
      (* Hinweis:
         - Quittierung der Scheibe
         - Uebergrosse Scheibe: Korrekturfahrt des Glastransports auf Anforderung des Greifers
      *)
      bprtScheibe := Greifer.bprtScheibe;

      tonlUeberwachungGreifer( IN := TRUE, PT := cZEIT_UEBERWACHUNG_GREIFER );

      IF ( Greifer.bpKorrekturfahrtAnfordern ) THEN
        Glastransport.bpKorrekturfahrtRueckwaerts := Greifer.bpKorrekturfahrtRueckwaerts;
        Glastransport.bpStarteKorrekturfahrt      := TRUE;
      ELSE
        Glastransport.bpStarteKorrekturfahrt      := FALSE;
      END_IF

      IF ( Greifer.bpEintransportAbgeschlossen ) THEN
        tonlUeberwachungGreifer( IN := FALSE );
        Greifer.bpStarteEintransport         := FALSE;
        Glastransport.bpStarteKorrekturfahrt := FALSE;
        steplAktion := STEP_1000_E;
      END_IF

      IF ( tonlUeberwachungGreifer.Q ) THEN
        tonlUeberwachungGreifer( IN := FALSE );
        Greifer.bpStarteEintransport         := FALSE;
        Glastransport.bpStarteKorrekturfahrt := FALSE;
        BasisStationsParameter.wFehlerNummer := cMELDUNG_GREIFER_STOESSEL_ABLAUF_ZEITUEBERSCHREITUNG;
        steplAktion := STEP_900_E;
      END_IF

    // EINTRANSPORT ==============================
    STEP_900_E:
      BasisStationsParameter.bFehler := TRUE;

    // EINTRANSPORT ==============================
    STEP_1000_E:
      bprtScheibe := FALSE;
      BasisStationsParameter.bEintransportAbgeschlossen[wWand] := TRUE;

  // EINTRANSPORT ==============================
  END_CASE
ELSE

  IF (steplAktion > STEP_0_E) THEN

    BasisStationsParameter.bEintransportAbgeschlossen[wWand] := FALSE;
    bprtScheibe := FALSE;

    Kippen.bpPositionieren := FALSE;
    Wandverstellung.bpStartePositionierung := FALSE;

    IF ( blMitGreifer ) THEN
      Greifer.bpStarteVorabPositionierungEintransport := FALSE;
      Greifer.bpStarteEintransport                    := FALSE;
      Glastransport.bpStarteKorrekturfahrt            := FALSE;
      tonlUeberwachungGreifer( IN := FALSE );
      blMitGreifer := FALSE;
    END_IF

    steplAktion := STEP_0_E;
  END_IF

END_IF
END_FUNCTION_BLOCK
